(* IEC 61131-3 sources: Versio-VersionControlSystem/fixtures/projects/TC3_PlcSample_reStrText/TC3_PlcSample_reStrText/LibraryDocumentationSample Project/LibPOUs/B_DocuElements/Hyperlinks/Footnotes, 5 files *)

(* ---- FB_Libdoc_AutomaticallyNumberedFootnotes.st ---- *)
(*

**Autonumbered footnotes**

Autonumbered footnotes are possible, like using [#]_ and [#]_.

--------

.. [#] This is the first one.

.. [#] This is the second one.
*)

FUNCTION_BLOCK FB_Libdoc_AutomaticallyNumberedFootnotes
VAR_INPUT
    nVarA : INT;
    nVarB : INT;
END_VAR
VAR_OUTPUT
    nSum : INT;
END_VAR
VAR
END_VAR

(* ---- FB_Libdoc_AutomaticallySymbolFootnotes.st ---- *)
(*

Here is a symbolic
footnote reference: [*]_ footnote reference: [*]_
footnote reference: [*]_ footnote reference: [*]_
footnote reference: [*]_ footnote reference: [*]_
footnote reference: [*]_ footnote reference: [*]_
footnote reference: [*]_ footnote reference: [*]_
footnote reference: [*]_

.. [*] This is the first footnote.
.. [*] This is the second footnote.
.. [*] This is the third footnote.
.. [*] This is the fourth footnote.
.. [*] This is the fifth footnote.
.. [*] This is the sixth footnote.
.. [*] This is the seventh footnote.
.. [*] This is the eighth footnote.
.. [*] This is the ninth footnote.
.. [*] This is the tenth footnote.
.. [*] This is the eleventh footnote.
*)

FUNCTION_BLOCK FB_Libdoc_AutomaticallySymbolFootnotes
VAR_INPUT
    nVarA : INT;
    nVarB : INT;
END_VAR
VAR_OUTPUT
    nSum : INT;
END_VAR
VAR
END_VAR

(* ---- FB_Libdoc_ManuallyAndAutomaticallyNumberedFootnotes.st ---- *)
(*

[2]_ will be "2" (manually numbered footnote),

[3]_ will be "3" (another manually numbered footnote),

[#]_ will be "4" (anonymous auto-numbered footnote), and

[#label]_ will be "1" (labeled auto-numbered).

--------

.. [2] This footnote is labeled manually, so its number is fixed.

.. [3] This footnote is also labeled manually, so its number is also fixed.

.. [#label] This autonumber-labeled footnote will be labeled "1".
   It is the first auto-numbered footnote and no other footnote
   with label "1" exists.  The order of the footnotes is used to
   determine numbering, not the order of the footnote references!

.. [#] This footnote will be labeled "4".  It is the second
   auto-numbered footnote, but footnote labels "1", "2", "3" are already used.
*)

FUNCTION_BLOCK FB_Libdoc_ManuallyAndAutomaticallyNumberedFootnotes
VAR_INPUT
    nVarA : INT;
    nVarB : INT;
END_VAR
VAR_OUTPUT
    nSum : INT;
END_VAR
VAR
END_VAR

(* ---- FB_Libdoc_ManuallyNumberedFootnotes.st ---- *)
(*

**Numerical footnote**

Footnote references, like [5]_. Note that footnotes may get rearranged, e.g., to the bottom of the "page".

--------

.. [5] A numerical footnote. Note there's no colon after the ``]``.
*)

FUNCTION_BLOCK FB_Libdoc_ManuallyNumberedFootnotes
VAR_INPUT
    nVarA : INT;
    nVarB : INT;
END_VAR
VAR_OUTPUT
    nSum : INT;
END_VAR
VAR
END_VAR

(* ---- FB_Libdoc_NamedAutomaticallyNumberedFootnotes.st ---- *)
(*

**Autonumbered labeled footnotes**

They may be assigned 'autonumber labels' - for instance, [#first]_ and [#second]_.

--------

.. [#first] a.k.a. first_

.. [#second] a.k.a. second_
*)

FUNCTION_BLOCK FB_Libdoc_NamedAutomaticallyNumberedFootnotes
VAR_INPUT
    nVarA : INT;
    nVarB : INT;
END_VAR
VAR_OUTPUT
    nSum : INT;
END_VAR
VAR
END_VAR
